Fanuc KAREL source: ks00031.KL

PROGRAM KS00031
%STACKSIZE=65535
%PRIORITY=65535
%NOLOCKGROUP
VAR
FLAG : BOOLEAN
N : INTEGER
STATUS : INTEGER
PN : STRING[80]
VN : STRING[80]
-- UNRESOLVED DECLARATIONS (source type spelling not recovered)
-- A : ARRAY[4] OF TYPE_0x001C (type_u16=0x201C)
-- B : ARRAY[4] OF TYPE_0x001C (type_u16=0x201C)
BEGIN
PN=''
VN='A'
-- UNRESOLVED_PC line 19 opcodes [22 22 1E] marker_code=27
END KS00031
